Staubli VAL3: forItem.dtx

public num nLoopValue
public bool bIOdisable
public string sIOindex
public string sForTRAJ
